(* IEC 61131-3 sources: codesys-to-s7/tests/corpus/C2S7-SEM-TIMER-Q/neg, 1 file *)

(* ---- input.st ---- *)
FUNCTION_BLOCK FB_Case
VAR
    tDelay : TON;
    x : BOOL;
    y : BOOL;
END_VAR
tDelay(IN := x, PT := T#1S);
y := tDelay.Q;
END_FUNCTION_BLOCK
